TYPE ST_PolarIIChamber_SupplyParam :
STRUCT
	Setpoint : DINT; // 1:1, ml/sec for liquid or Pa for gas
END_STRUCT
END_TYPE

(* stored: Version 1.1.0.1, ProductVersion 3.1.4026.18
   DUT ST_PolarIIChamber_SupplyParam: Id {14000000-0000-0000-0000-000000000013} *)
